Fanuc KAREL source: KD00059.KL

PROGRAM KD00059
%NOLOCKGROUP
VAR
  I: INTEGER
  J: INTEGER
  B: BOOLEAN
  R: REAL
  S: STRING[80]
BEGIN
  CONDITION[1]:
  WHEN DIN[1] = ON DO
    CANCEL
  ENDCONDITION
END KD00059
